(* PLC project Unnamed, Unknown Unnamed 1 *)
(* stored: creationDateTime 2026-09-08T11:20:29, modificationDateTime 2026-09-08T11:20:29 *)

FUNCTION_BLOCK TOF
  VAR_OUTPUT
    Q : BOOL;
    ET : TIME;
  END_VAR
  VAR_INPUT
    IN : BOOL;
    PT : TIME;
  END_VAR

END_FUNCTION_BLOCK

PROGRAM main
  VAR
    stop : BOOL;
    start : BOOL;
    machine_run : BOOL;
    TOF0 : TOF;
    fan : BOOL;
  END_VAR

(* LD diagram, written out as Structured Text *)
machine_run := NOT stop AND (start OR machine_run);
fan := TOF0.Q;
TOF0(IN := machine_run, PT := T#10s);
END_PROGRAM

CONFIGURATION Config0
  RESOURCE Res0 ON PLC
    TASK task0(INTERVAL := T#20ms, PRIORITY := 1);
    PROGRAM instance0 WITH task0 : main;
  END_RESOURCE
END_CONFIGURATION
